(* IEC 61131-3 sources: plc-process-lib/tests/POUs/Suites/FB_Pid_Test (part 2) *)

(* ---- SpTrackPvManualSetpointFollowsPv.method.decl.st ---- *)
// xSpTrackPv: в Manual задание следует за PV (ФБ пишет PV в stCmd.rSp_eu), поэтому переход в
// Auto идёт с нулевой ошибкой и выход не меняется.
METHOD PRIVATE SpTrackPvManualSetpointFollowsPv
VAR
    fbTime   : FB_FakeTime;       // подменное время, старт 1 ч
    fbPid    : FB_PID;            // ФБ под тестом
    stCmd    : ST_PidCmd;         // команды
    stRetain : ST_DeviceRetain;   // режим: старт в Manual
    stCfg    : ST_PidCfg;         // конфигурация теста
    iStep    : INT;               // шаг цикла
    rCmdSp   : REAL;              // stCmd.rSp_eu в Manual
    rOutSw   : REAL;              // выход в вызове перехода
END_VAR

(* ---- SpTrackPvManualSetpointFollowsPv.method.impl.st ---- *)
coUnit.TEST('Pid_SpTrackPv_ManualSetpoint_FollowsPv');
// источник: tools/reference/pid.py, сценарий sp_track_pv
stCfg.rKp := 2.0;
stCfg.rTi_s := 10.0;
stCfg.xSpTrackPv := TRUE;
stCmd.rManualOut_pct := 30.0;
stCmd.rSp_eu := 50.0;
fbPid.rPv_eu := 47.5;
fbPid.xPvValid := TRUE;
fbPid(itfTime := fbTime, stCmd := stCmd, stRetain := stRetain, stCfg := stCfg);       // t0: Manual
FOR iStep := 1 TO 5 DO
    fbTime.Advance(tStep := T#100MS);
    fbPid(itfTime := fbTime, stCmd := stCmd, stRetain := stRetain, stCfg := stCfg);
END_FOR
rCmdSp := stCmd.rSp_eu;
fbTime.Advance(tStep := T#100MS);
stCmd.stCommon.xSetAuto := TRUE;
fbPid(itfTime := fbTime, stCmd := stCmd, stRetain := stRetain, stCfg := stCfg);       // Manual -> Auto
rOutSw := fbPid.rOut_pct;
FOR iStep := 1 TO 10 DO
    fbTime.Advance(tStep := T#100MS);
    fbPid(itfTime := fbTime, stCmd := stCmd, stRetain := stRetain, stCfg := stCfg);
END_FOR
// ref: sp_track_pv.cmd_sp
AssertEquals_REAL(Expected := 47.5, Actual := rCmdSp, Delta := 0.0, Message := 'SP follows PV in Manual');
// ref: sp_track_pv.out_switch
AssertEquals_REAL(Expected := 30.0, Actual := rOutSw, Delta := 1.0E-4, Message := 'no bump at Manual -> Auto');
// ref: sp_track_pv.out_1s
AssertEquals_REAL(Expected := 30.0, Actual := fbPid.rOut_pct, Delta := 1.0E-4, Message := 'zero error after switch');
AssertEquals_REAL(Expected := 47.5, Actual := stCmd.rSp_eu, Delta := 0.0, Message := 'SP no longer written in Auto');
coUnit.TEST_FINISHED();

(* ---- StartupOutActInitialisesOutput.method.decl.st ---- *)
// Старт ПЛК в Auto (режим из stRetain) с xUseOutAct: stCmd.rManualOut_pct = 0 (GVL_Hmi после
// потери питания не сохраняется), механизм стоит на 37 % — выход первого вызова берётся из
// rOutAct_pct, интегратор инициализируется под него (I = 37 - 8 = 29 %), и регулирование идёт от
// 37 % без провала в ноль. Второй экземпляр: rOutAct_pct не конечен — выход из rManualOut_pct.
METHOD PRIVATE StartupOutActInitialisesOutput
VAR
    fbTime    : FB_FakeTime;       // подменное время, старт 1 ч
    fbPid     : FB_PID;            // ФБ под тестом: rOutAct_pct = 37 %
    fbPidNaN  : FB_PID;            // второй экземпляр: rOutAct_pct не конечен
    stCmd     : ST_PidCmd;         // команды: rManualOut_pct = 0
    stCmdNaN  : ST_PidCmd;         // команды второго экземпляра: rManualOut_pct = 42 %
    stRetain  : ST_DeviceRetain;   // режим Auto из Persistent Variables
    stRetNaN  : ST_DeviceRetain;   // то же для второго экземпляра
    stCfg     : ST_PidCfg;         // конфигурация теста
    uBits     : U_RealBits;        // источник NaN
    iStep     : INT;               // шаг цикла
    rOutSt    : REAL;              // выход первого вызова
    rISt      : REAL;              // интегратор первого вызова
    rCmdOutSt : REAL;              // stCmd.rManualOut_pct после первого вызова
END_VAR

(* ---- StartupOutActInitialisesOutput.method.impl.st ---- *)
coUnit.TEST('Pid_Startup_OutActInitialisesOutput');
// источник: tools/reference/pid.py, сценарий start_outact
uBits.dwValue := 16#7FC00000;                                                          // тихий NaN
stCfg.rKp := 2.0;
stCfg.rTi_s := 10.0;
stCfg.xUseOutAct := TRUE;
stRetain.eRemoteMode := E_DeviceMode.Auto;
stRetNaN := stRetain;
stCmd.rSp_eu := 50.0;
stCmdNaN := stCmd;
stCmdNaN.rManualOut_pct := 42.0;
fbPid.rPv_eu := 46.0;                                                                  // e = 4 %, P = 8 %
fbPid.xPvValid := TRUE;
fbPid.rOutAct_pct := 37.0;                                                             // механизм на 37 %
fbPidNaN.rPv_eu := 46.0;
fbPidNaN.xPvValid := TRUE;
fbPidNaN.rOutAct_pct := uBits.rValue;
fbPid(itfTime := fbTime, stCmd := stCmd, stRetain := stRetain, stCfg := stCfg);       // первый вызов
fbPidNaN(itfTime := fbTime, stCmd := stCmdNaN, stRetain := stRetNaN, stCfg := stCfg);
rOutSt := fbPid.rOut_pct;
rISt := fbPid.stSts.rI_pct;
rCmdOutSt := stCmd.rManualOut_pct;
FOR iStep := 1 TO 2 DO                                                                 // механизм отрабатывает выход
    fbPid.rOutAct_pct := fbPid.rOut_pct;
    fbTime.Advance(tStep := T#100MS);
    fbPid(itfTime := fbTime, stCmd := stCmd, stRetain := stRetain, stCfg := stCfg);
END_FOR
AssertTrue(Condition := fbPid.Mode = E_DeviceMode.Auto, Message := 'Auto restored from retain');
// ref: start_outact.out_start
AssertEquals_REAL(Expected := 37.0, Actual := rOutSt, Delta := 1.0E-4, Message := 'output from rOutAct_pct, not 0');
// ref: start_outact.i_start
AssertEquals_REAL(Expected := 29.0, Actual := rISt, Delta := 1.0E-4, Message := 'I = u - P at startup');
AssertEquals_REAL(Expected := 37.0, Actual := rCmdOutSt, Delta := 0.0,
                  Message := 'rManualOut_pct tracks startup output');
// ref: start_outact.out_2
AssertEquals_REAL(Expected := 37.08, Actual := fbPid.rOut_pct, Delta := 1.0E-4, Message := 'control continues from 37');
// AssertEquals_REAL пропускает NaN (ABS(NaN) > Delta = FALSE): конечность проверяется отдельно
AssertTrue(Condition := F_IsFinite(rIn := fbPidNaN.rOut_pct), Message := 'NaN source: output stays finite');
// ref: start_outact.out_start_nan
AssertEquals_REAL(Expected := 42.0, Actual := fbPidNaN.rOut_pct, Delta := 1.0E-4,
                  Message := 'non-finite rOutAct_pct: output from rManualOut_pct');
coUnit.TEST_FINISHED();

(* ---- TimeBackwardsInitStepNoJump.method.decl.st ---- *)
// «Время назад» на 30 с (источник времени переставлен): LTIME без знака, разность не считается;
// шаг инициализации — выход прежний, бит DT_GAP; дальше интегрирование по обычному шагу.
METHOD PRIVATE TimeBackwardsInitStepNoJump
VAR
    fbTime   : FB_FakeTime;       // подменное время, старт 1 ч
    fbPid    : FB_PID;            // ФБ под тестом
    stCmd    : ST_PidCmd;         // команды
    stRetain : ST_DeviceRetain;   // режим: старт в Manual
    stCfg    : ST_PidCfg;         // конфигурация теста
    iStep    : INT;               // шаг цикла
    rBefore  : REAL;              // выход до скачка времени
    rBack    : REAL;              // выход в вызове после скачка
    wStsBack : WORD;              // wStatus в вызове после скачка
    rAfter   : REAL;              // выход в следующем вызове
END_VAR

(* ---- TimeBackwardsInitStepNoJump.method.impl.st ---- *)
coUnit.TEST('Pid_TimeBackwards_InitStep_NoJump');
// источник: tools/reference/pid.py, сценарий time_back
stCfg.rKp := 2.0;
stCfg.rTi_s := 10.0;
stCmd.rManualOut_pct := 30.0;
stCmd.rSp_eu := 50.0;
fbPid.rPv_eu := 50.0;
fbPid.xPvValid := TRUE;
fbPid(itfTime := fbTime, stCmd := stCmd, stRetain := stRetain, stCfg := stCfg);       // t0: Manual
fbTime.Advance(tStep := T#100MS);
stCmd.stCommon.xSetAuto := TRUE;
fbPid(itfTime := fbTime, stCmd := stCmd, stRetain := stRetain, stCfg := stCfg);       // Auto
fbPid.rPv_eu := 46.0;                                                                  // e = 4 %
FOR iStep := 1 TO 10 DO
    fbTime.Advance(tStep := T#100MS);
    fbPid(itfTime := fbTime, stCmd := stCmd, stRetain := stRetain, stCfg := stCfg);
END_FOR
rBefore := fbPid.rOut_pct;
fbTime.SetNow(ltValue := fbTime.Now() - LTIME#30S);                                    // время назад
fbPid(itfTime := fbTime, stCmd := stCmd, stRetain := stRetain, stCfg := stCfg);
rBack := fbPid.rOut_pct;
wStsBack := fbPid.stSts.stCommon.wStatus;
fbTime.Advance(tStep := T#100MS);
fbPid(itfTime := fbTime, stCmd := stCmd, stRetain := stRetain, stCfg := stCfg);
rAfter := fbPid.rOut_pct;
fbTime.Advance(tStep := T#100MS);
fbPid(itfTime := fbTime, stCmd := stCmd, stRetain := stRetain, stCfg := stCfg);
// ref: time_back.out_before
AssertEquals_REAL(Expected := 38.72, Actual := rBefore, Delta := 1.0E-4, Message := 'output before time jump');
// ref: time_back.out_back
AssertEquals_REAL(Expected := 38.72, Actual := rBack, Delta := 1.0E-4, Message := 'time backwards: output held');
AssertEquals_WORD(Expected := GVL_Const.PID_STS_DT_GAP, Actual := wStsBack AND GVL_Const.PID_STS_DT_GAP,
                  Message := 'status bit DT_GAP');
// ref: time_back.out_after
AssertEquals_REAL(Expected := 38.72, Actual := rAfter, Delta := 1.0E-4, Message := 'first normal step');
// ref: time_back.out_after2
AssertEquals_REAL(Expected := 38.8, Actual := fbPid.rOut_pct, Delta := 1.0E-4, Message := 'integration resumes');
coUnit.TEST_FINISHED();

(* ---- TrackNaNValueHoldsOutput.method.decl.st ---- *)
// Слежение за неконечным значением (NaN из образа обмена): выход и слежение в Cmd остаются
// прежними, NaN на механизм не уходит; конечное значение снова принимается.
METHOD PRIVATE TrackNaNValueHoldsOutput
VAR
    fbTime   : FB_FakeTime;       // подменное время, старт 1 ч
    fbPid    : FB_PID;            // ФБ под тестом
    stCmd    : ST_PidCmd;         // команды
    stRetain : ST_DeviceRetain;   // режим
    stCfg    : ST_PidCfg;         // конфигурация теста
    uBits    : U_RealBits;        // источник NaN
    rOutNaN  : REAL;              // выход при NaN
    rCmdNaN  : REAL;              // stCmd.rManualOut_pct при NaN
END_VAR

(* ---- TrackPresetsIntegratorBumplessRelease.method.decl.st ---- *)
// Слежение в Auto (Kp = 2, Ti = 10 с, нижний предел 10 %): выход = rTrack_pct без пределов (0 %),
// интегратор I = u - P - D, бит TRACKING, Cmd следит за выходом; после снятия xTrack выход
// продолжается с 25 % без рывка. Available = FALSE при слежении (PV годна, Auto), TRUE после снятия.
METHOD PRIVATE TrackPresetsIntegratorBumplessRelease
VAR
    fbTime    : FB_FakeTime;       // подменное время, старт 1 ч
    fbPid     : FB_PID;            // ФБ под тестом
    stCmd     : ST_PidCmd;         // команды
    stRetain  : ST_DeviceRetain;   // режим: Auto из Retain
    stCfg     : ST_PidCfg;         // конфигурация теста
    iStep     : INT;               // шаг цикла
    rOutTrk0  : REAL;              // выход при слежении за 0 %
    xTrkBit0  : BOOL;              // бит TRACKING при слежении
    rOutRel   : REAL;              // выход в вызове снятия слежения
END_VAR

(* ---- TrackPresetsIntegratorBumplessRelease.method.impl.st ---- *)
coUnit.TEST('Pid_Track_PresetsIntegrator_BumplessRelease');
// источник: tools/reference/pid.py, сценарий track
stCfg.rKp := 2.0;
stCfg.rTi_s := 10.0;
stCfg.rOutMin_pct := 10.0;
stCfg.rSafeOut_pct := 10.0;                                                            // в пределах выхода (бит 11)
stRetain.eRemoteMode := E_DeviceMode.Auto;
stCmd.rSp_eu := 50.0;
fbPid.rPv_eu := 47.0;                                                                  // e = 3 %, P = 6
fbPid.xPvValid := TRUE;
fbPid.xTrack := TRUE;
fbPid.rTrack_pct := 0.0;                                                               // механизм стоит
fbPid(itfTime := fbTime, stCmd := stCmd, stRetain := stRetain, stCfg := stCfg);       // t0: Auto, слежение
rOutTrk0 := fbPid.rOut_pct;
xTrkBit0 := (fbPid.stSts.stCommon.wStatus AND GVL_Const.PID_STS_TRACKING) <> 0;
fbPid.rTrack_pct := 25.0;
FOR iStep := 1 TO 10 DO
    fbTime.Advance(tStep := T#100MS);
    fbPid(itfTime := fbTime, stCmd := stCmd, stRetain := stRetain, stCfg := stCfg);
END_FOR
// ref: track.out_track0
AssertEquals_REAL(Expected := 0.0, Actual := rOutTrk0, Delta := 1.0E-4, Message := 'tracking ignores rOutMin_pct');
AssertTrue(Condition := xTrkBit0, Message := 'status bit TRACKING');
// ref: track.out_track
AssertEquals_REAL(Expected := 25.0, Actual := fbPid.rOut_pct, Delta := 1.0E-4, Message := 'output = rTrack_pct');
// ref: track.i_track
AssertEquals_REAL(Expected := 19.0, Actual := fbPid.stSts.rI_pct, Delta := 1.0E-4, Message := 'I preset = 25 - 6');
AssertEquals_REAL(Expected := 25.0, Actual := stCmd.rManualOut_pct, Delta := 1.0E-4, Message := 'Cmd tracks output');
AssertFalse(Condition := fbPid.Available, Message := 'not available while tracking, PV valid in Auto');
fbPid.xTrack := FALSE;
fbTime.Advance(tStep := T#100MS);
fbPid(itfTime := fbTime, stCmd := stCmd, stRetain := stRetain, stCfg := stCfg);       // слежение снято
rOutRel := fbPid.rOut_pct;
FOR iStep := 1 TO 10 DO
    fbTime.Advance(tStep := T#100MS);
    fbPid(itfTime := fbTime, stCmd := stCmd, stRetain := stRetain, stCfg := stCfg);
END_FOR
// ref: track.out_release
AssertEquals_REAL(Expected := 25.0, Actual := rOutRel, Delta := 1.0E-4, Message := 'no bump at release');
// ref: track.out_release_1s
AssertEquals_REAL(Expected := 25.6, Actual := fbPid.rOut_pct, Delta := 1.0E-4, Message := 'then integral action');
AssertEquals_WORD(Expected := 0, Actual := fbPid.stSts.stCommon.wStatus AND GVL_Const.PID_STS_TRACKING,
                  Message := 'TRACKING cleared');
AssertTrue(Condition := fbPid.Available, Message := 'available after release');
coUnit.TEST_FINISHED();

(* ---- TrackPvMovingNoDerivativeKickAtRelease.method.decl.st ---- *)
// Слежение при движущейся PV и Td > 0: D работает и при слежении (за 2 с выходит на 5 %), а
// предустановка I := u - P - D держит v = u. Снятие слежения — выход 30 % плюс изменение P и D за
// один шаг, без «удара» на величину D.
METHOD PRIVATE TrackPvMovingNoDerivativeKickAtRelease
VAR
    fbTime   : FB_FakeTime;       // подменное время, старт 1 ч
    fbPid    : FB_PID;            // ФБ под тестом
    stCmd    : ST_PidCmd;         // команды
    stRetain : ST_DeviceRetain;   // режим: Auto из Retain
    stCfg    : ST_PidCfg;         // конфигурация теста
    iStep    : INT;               // шаг цикла
    rDTrk    : REAL;              // D в конце слежения
    rITrk    : REAL;              // I в конце слежения
    rOutTrk  : REAL;              // выход в конце слежения
END_VAR

(* ---- TrackPvMovingNoDerivativeKickAtRelease.method.impl.st ---- *)
coUnit.TEST('Pid_Track_PvMoving_NoDerivativeKickAtRelease');
// источник: tools/reference/pid.py, сценарий track_d
stCfg.rKp := 2.0;
stCfg.rTi_s := 10.0;
stCfg.rTd_s := 1.0;                                                                    // N = 10: Tf = 0,1 с
stRetain.eRemoteMode := E_DeviceMode.Auto;
stCmd.rSp_eu := 50.0;
fbPid.rPv_eu := 50.0;
fbPid.xPvValid := TRUE;
fbPid.xTrack := TRUE;
fbPid.rTrack_pct := 30.0;
fbPid(itfTime := fbTime, stCmd := stCmd, stRetain := stRetain, stCfg := stCfg);       // t0: Auto, слежение
FOR iStep := 1 TO 20 DO                                                                // 2 с, PV падает 2,5 %/с
    fbPid.rPv_eu := fbPid.rPv_eu - 0.25;
    fbTime.Advance(tStep := T#100MS);
    fbPid(itfTime := fbTime, stCmd := stCmd, stRetain := stRetain, stCfg := stCfg);
END_FOR
rDTrk := fbPid.stSts.rD_pct;
rITrk := fbPid.stSts.rI_pct;
rOutTrk := fbPid.rOut_pct;
fbPid.xTrack := FALSE;                                                                 // слежение снято
fbPid.rPv_eu := fbPid.rPv_eu - 0.25;
fbTime.Advance(tStep := T#100MS);
fbPid(itfTime := fbTime, stCmd := stCmd, stRetain := stRetain, stCfg := stCfg);
// ref: track_d.d_track
AssertEquals_REAL(Expected := 4.999995, Actual := rDTrk, Delta := 1.0E-4, Message := 'D works while tracking');
// ref: track_d.i_track
AssertEquals_REAL(Expected := 15.000005, Actual := rITrk, Delta := 1.0E-4, Message := 'I preset = u - P - D');
// ref: track_d.out_track
AssertEquals_REAL(Expected := 30.0, Actual := rOutTrk, Delta := 1.0E-4, Message := 'output = rTrack_pct');
// ref: track_d.out_release
AssertEquals_REAL(Expected := 30.500002, Actual := fbPid.rOut_pct, Delta := 1.0E-4,
                  Message := 'release: one-step change of P and D only, no derivative kick');
// ref: track_d.d_release
AssertEquals_REAL(Expected := 4.999998, Actual := fbPid.stSts.rD_pct, Delta := 1.0E-4, Message := 'D continues');
coUnit.TEST_FINISHED();

(* ---- TrackWithInvalidPvNoFailure.method.decl.st ---- *)
// Слежение в Auto при негодной PV: ПИД не регулирует, поэтому не Failure и wFault = 0; выход —
// rTrack_pct; тревога PvInvalid по контракту (PV негодна в Auto) активна.
METHOD PRIVATE TrackWithInvalidPvNoFailure
VAR
    fbTime   : FB_FakeTime;       // подменное время, старт 1 ч
    fbPid    : FB_PID;            // ФБ под тестом
    stCmd    : ST_PidCmd;         // команды
    stRetain : ST_DeviceRetain;   // режим: Auto из Retain
    stCfg    : ST_PidCfg;         // конфигурация по умолчанию
END_VAR
